// TIA Portal V21 export
// export: Created 2026-08-21T20:18:51.8529801Z, ExportSetting None, DisplayName Totally Integrated Automation Portal, DisplayVersion V21, DisplayName STEP 7 Professional, DisplayVersion V21, DisplayName STEP 7 Safety, DisplayVersion V21, DisplayName Tech WebApplication, DisplayVersion V21, DisplayName WinCC Basic/Comfort/Advanced, DisplayVersion V21, DisplayName WinCC Professional, DisplayVersion V21, DisplayName WinCC Unified, DisplayVersion V21
DATA_BLOCK "LAH100_Type"   // DB19
// stored: InstanceOfName MTPBinMon_Type1, InstanceOfType FB
"MTPBinMon_Type1"
   // VAR_INPUT
   //    PV { ExternalAccessible := 'False'; ExternalVisible := 'False'; ExternalWritable := 'False'} : Bool;
   //    PV_QB { ExternalAccessible := 'False'; ExternalVisible := 'False'; ExternalWritable := 'False'} : Bool;
   //    InvPV_In { ExternalAccessible := 'False'; ExternalVisible := 'False'; ExternalWritable := 'False'} : Bool;
   // END_VAR
   // VAR_OUTPUT
   //    PV_Out { ExternalAccessible := 'False'; ExternalVisible := 'False'; ExternalWritable := 'False'} : Bool;
   //    to_Indicate { ExternalAccessible := 'False'; ExternalVisible := 'False'; ExternalWritable := 'False'} : "StruCm";
   // END_VAR
   // VAR
   //    DiIn_IDB { ExternalAccessible := 'False'; ExternalVisible := 'False'; ExternalWritable := 'False'} : "DiIn";
   //    MonDiL_IDB { S7_SetPoint := 'True'} : "MonDiL";
   //    MTPBinMon_IDB { ExternalVisible := 'False'; S7_SetPoint := 'True'} : "MTPBinMon";
   // END_VAR
BEGIN
END_DATA_BLOCK
